TYPE ST_EL3356ChannelCtrl_1 :
STRUCT
	bStartCalibration			:BOOL;			(* Ctrl start calibration *)
	bDisableCalibration		:BOOL;			(* Ctrl disable calibration *)
	bInputFreeze				:BOOL;			(* Ctrl input freeze *)
	bTare					:BOOL;			(* Ctrl tare *)
END_STRUCT
END_TYPE

(* stored: Version 1.1.0.1, ProductVersion 3.1.4024.15
   DUT ST_EL3356ChannelCtrl_1: Id {07aca0fb-67c5-4421-b247-656463332a1f} *)
